// Mitsubishi GX Works2 project: AVRInfacomV3   PLC: FX3G

TYPE CutCard : STRUCT
  Lenth : DINT;
  Qnt : DINT;
END_STRUCT END_TYPE

// global labels: _io
VAR_GLOBAL
  DI_Avar1 AT X000 : BOOL;
  DI_Line1IsOff AT X001 : BOOL;
  DI_Avar2 AT X002 : BOOL;
  DI_Line2IsOff AT X003 : BOOL;
  DI_AvarGenerator AT X004 : BOOL;
  DI_GeneratorIsOff AT X005 : BOOL;
  DI_AvarSection AT X006 : BOOL;
  DI_SectionIsOff AT X007 : BOOL;
  DI_RKF1 AT X010 : BOOL;
  DI_RKF2 AT X011 : BOOL;
  DI_RKF3 AT X012 : BOOL;
  DI_Avarkontrol AT X013 : BOOL;
  DO_On1 AT Y000 : BOOL;
  DO_Off1 AT Y001 : BOOL;
  DO_On2 AT Y002 : BOOL;
  DO_Off2 AT Y003 : BOOL;
  DO_OnGenerator AT Y004 : BOOL;
  DO_OffGenerator AT Y005 : BOOL;
  DO_OnSection AT Y006 : BOOL;
  DO_OffSection AT Y007 : BOOL;
  DO_StartGenerator AT Y010 : BOOL;
END_VAR

// global labels: _gvl
VAR_GLOBAL
  gxAvto AT M400 : BOOL;
  gxOn1 AT M100 : BOOL;
  gxOff1 AT M101 : BOOL;
  gxOn2 AT M102 : BOOL;
  clTimeGenerator AT D1000 : INT;
  clTimeRKF1 AT D1001 : INT;
  clTimeRKF2 AT D1002 : INT;
  clTimeRKF3 AT D1003 : INT;
  gxOff2 AT M103 : BOOL;
  gxOnGenerator AT M104 : BOOL;
  gxOffGenerator AT M105 : BOOL;
  gxOnSection AT M106 : BOOL;
  gxOffSection AT M107 : BOOL;
  gxStartGenerator AT M108 : BOOL;
  clStartgenerator AT D1004 : INT;
  gxIsAlarm AT M150 : BOOL;
  VVALine1 : VVA;
  VVALine2 : VVA;
  VVAGen : VVA;
  VVASec : VVA;
  clTimeBackAuto AT D1005 : INT;
  gxVVAOff AT M401 : BOOL;
  gxProblemVVA1 AT M110 : BOOL;
  gxProblemVVA2 AT M111 : BOOL;
  gxProblemVVAgen AT M112 : BOOL;
END_VAR

// task Task_init (event M8002, interval 0, priority 1): PRG_INIT
// task Task_Main (event TRUE, interval 0, priority 31): POU_01
// task Task_Process (event TRUE, interval 0, priority 31): PRG_PROCESS
// user libraries (not included): AlarmManger128, Modbusv16, TimeControl, Utils

PROGRAM POU_01
VAR
  fbAmBlock : AM_IS_BLOCK;
  iStep : INT;
  wTimeRKFs : INT;
  xGenerator : BOOL;
  TPStartGen : TP;
  fbAmalarm : AM_HAS_ALARMS;
  xAllGood : BOOL;
END_VAR
(* fbAmBlock(iProcessNum := 1, iSeverity := AM_ERROR, Q := gxIsAlarm); *)
fbAmalarm(iProcessNum := 0, iSeverity := 0, Q := gxIsAlarm);
wTimeRKFs := SEL(clTimeRKF1 > clTimeRKF2, clTimeRKF2, clTimeRKF1);

IF MEF(gxAvto) THEN
    iStep := 10;
END_IF;

IF MEP(gxAvto) THEN
    iStep := 0;
END_IF;

M1 := DI_RKF1 AND NOT VVALine1.xError;
M2 := DI_RKF2 AND NOT VVALine2.xError;
M3 := DI_RKF3 AND NOT VVAGen.xError;

OUT_T(M1, TC1, SEC_TO_TIMER100(clTimeRKF1));
OUT_T(M2, TC2, SEC_TO_TIMER100(clTimeRKF2));
OUT_T(M3, TC3, SEC_TO_TIMER100(clTimeRKF3)); 

OUT_T(TRUE, TC30, 100);
OUT_T(iStep = 30 AND DI_Line1IsOff, TC4, 100);
OUT_T(iStep = 40 AND DI_Line2IsOff, TC5, 100);
OUT_T(iStep = 50 AND DI_GeneratorIsOff, TC6, 100);

(*BackAuto
OUT_T(gxVVAOff, TC31, SEC_TO_TIMER100(clTimeBackAuto));
IF TS31 THEN
	gxVVAOff := FALSE;
END_IF;
*)

CASE iStep OF
    0: (* Reset timers *)
        xGenerator := FALSE;
        gxStartGenerator := FALSE;
        MOV(TS30, 1, iStep);

    1: (* Test everything *)
    	xAllGood := TRUE;
    	
    
        MOV(xAllGood, 10, iStep);

    10: (* Idle *)

        MOV(gxAvto, 20, iStep);
        RST(gxAvto, gxStartGenerator);

		SET(
			MEP(gxOn1) 
			AND DI_Line2IsOff 
			AND DI_Line1IsOff 
			AND DI_GeneratorIsOff 
			AND DI_RKF1, 
			VVALine1.SetOn
		);
		RST( 
			MEP(gxOff1) 
			OR NOT DI_Line2IsOff 
			OR NOT DI_GeneratorIsOff 
			OR NOT DI_RKF1, 
			VVALine1.SetOn
		);

		SET(
			MEP(gxOn2) 
			AND DI_Line2IsOff 
			AND DI_Line1IsOff 
			AND DI_GeneratorIsOff 
			AND DI_RKF2, 
			VVALine2.SetOn
		);
		RST( 
			MEP(gxOff2) 
			OR NOT DI_Line1IsOff 
			OR NOT DI_GeneratorIsOff 
			OR NOT DI_RKF2, 
			VVALine2.SetOn
		);
		
		SET(
			MEP(gxOnGenerator) 
			AND DI_Line2IsOff 
			AND DI_Line1IsOff 
			AND DI_GeneratorIsOff 
			AND DI_RKF3, 
			VVAGen.SetOn
		);
		RST( 
			MEP(gxOffGenerator) 
			OR NOT DI_Line1IsOff 
			OR NOT DI_Line2IsOff 
			OR NOT DI_RKF3, 
			VVAGen.SetOn
		);
      
        xGenerator := gxStartGenerator;

    20: (* Selector *)
        MOV(TS1, 30, iStep);
        MOV(TS2 AND NOT TS1, 40, iStep);
        MOV(NOT TS1 AND NOT TS2 AND TS3, 50, iStep);
		xGenerator := NOT TS1 AND NOT TS2;

    30: (* Line 1 *)
	    VVALine2.SetOn := FALSE;
	    VVAGen.SetOn := FALSE;
        SET(TS4, gxProblemVVA1);
        SET(TS4, gxVVAOff);
        
        MOV(
        	NOT TS1 (* Контроль фаз *)
        	OR TS4 (* выключение в ручну *)
        	OR VVALine1.xError, (* автомат в ошибке *)
        	10,
        	iStep
        );

        VVALine1.SetOn := DI_GeneratorIsOff 
        	AND DI_Line2IsOff AND iStep = 30;
    
    40: (* Line 2 *)
	    VVALine1.SetOn := FALSE;
	    VVAGen.SetOn := FALSE;
        SET(TS5, gxProblemVVA2);
        SET(TS5, gxVVAOff);
         
        MOV(
        	NOT TS2 (* Контроль фаз *)
        	OR TS5 (* выключение в ручну *)
        	OR VVALine2.xError, (* автомат в ошибке *)
        	10,
        	iStep
        );

        VVALine2.SetOn := DI_GeneratorIsOff 
        	AND DI_Line1IsOff AND iStep = 40;
    
    50: (* Generator *)
	    VVALine2.SetOn := FALSE;
	    VVALine1.SetOn := FALSE;
        SET(TS6, gxProblemVVAgen);
        SET(TS6, gxVVAOff);
        
        MOV(
        	NOT TS3 (* Контроль фаз *)
        	OR TS1 OR TS2 (* появилась сеть *)
        	OR TS6 (* выключение в ручну *)
        	OR VVAGen.xError, (* автомат в ошибке *)
        	10,
        	iStep
        );
		
		xGenerator := TRUE;
        VVAGen.SetOn := DI_Line1IsOff 
        	AND DI_Line2IsOff AND iStep = 50;
END_CASE;

TPStartGen(IN := xGenerator, PT := SEC_TO_TIME(clTimeGenerator));
DO_StartGenerator := NOT (xGenerator OR TPStartGen.Q);

IF iStep > 0 THEN
	VVALine1(
		IsOn := NOT DI_Line1IsOff, 
		ResetAlarm := M2002, 
		Vkl := DO_On1, 
		Otkl := DO_Off1
	);
	VVALine2(
		IsOn := NOT DI_Line2IsOff, 
		ResetAlarm := M2002, 
		Vkl := DO_On2, 
		Otkl := DO_Off2
	);
	VVAGen(
		IsOn := NOT DI_GeneratorIsOff, 
		ResetAlarm := M2002, 
		Vkl := DO_OnGenerator, 
		Otkl := DO_OffGenerator
	);
END_IF;
END_PROGRAM

PROGRAM PRG_INIT
VAR
  fbAmInit : AM_INIT;
END_VAR
AM_D_START := 3000;

VVALine1.AlarmNum := 1;
VVALine2.AlarmNum := 2;
VVAGen.AlarmNum := 3;
VVASec.AlarmNum := 4;

(* Ошибка UPS *)
fbAmInit(iNum := 0, iSeverity := 3, iProcess := 1, xLatch := 0, xBuzzer := 0, xLock := 0);
(* Ошибка ВА Сеть 1 *)
fbAmInit(iNum := 1 , xLatch := 1, xLock := 0 );
(* Ошибка ВА Сеть 2 *)
fbAmInit(iNum := 2 , xLatch := 1, xLock := 0 );
(* Ошибка ВА Генератор *)
fbAmInit(iNum := 3 , xLatch := 1, xLock := 0 );
(* Ошибка ВА Секционный *)
fbAmInit(iNum := 4 , xLatch := 1, xLock := 0);
(* Отказ вкл ВА Сеть 1 *)
fbAmInit(iNum := 5, xLatch := 0, xLock := 0);
(* Отказ выкл ВА Сеть 1 *)
fbAmInit(iNum := 6 , xLatch := 0, xLock := 0 );
(* Отказ вкл ВА Сеть 2 *)
fbAmInit(iNum := 7 , xLatch := 0, xLock := 0 );
(* Отказ выкл ВА Сеть 2 *)
fbAmInit(iNum := 8 , xLatch := 0, xLock := 0 );
(* Отказ вкл ВА Генератор *)
fbAmInit(iNum := 9 , xLatch := 0, xLock := 0);
(* Отказ выкл ВА Генератор *)
fbAmInit(iNum := 10, xLatch := 0, xLock := 0);
(* Отказ вкл ВА Секционный *)
fbAmInit(iNum := 11 , xLatch := 0, xLock := 0 );
(* Отказ выкл ВА Секционный *)
fbAmInit(iNum := 12 , xLatch := 0, xLock := 0 );
(* Отказ запуска генератора *)
fbAmInit(iNum := 13 , xLatch := 1, xLock := 0 );
(* Данные не заполнены *)
fbAmInit(iNum := 14 , xLatch := 0, xLock := 1);
END_PROGRAM

PROGRAM PRG_PROCESS
VAR
  fbAmSet : AM_SET;
  fbAmReset : AM_RST;
  xNodata : BOOL;
  fbAMEvents : AM_EVENT;
  fbTOFResetProblems : TOF;
  PortSettings : DWORD;
  xMBInit : BOOL;
END_VAR
fbAmReset(IN := M2002);

IF  M2002 THEN
	gxProblemVVA1 := FALSE;
	gxProblemVVA2 := FALSE;
	gxProblemVVAgen := FALSE;
END_IF;

PortSettings := MB_PORT_SETTINGS(MB_PARITY_NONE, MB_STOPBIT_1, MB_BPS_38400);
xMBInit :=  MB_SLAVE_INIT_PORT2(TRUE, 20, PortSettings);

(* Тревоги *)
OUT_T(NOT DI_Avarkontrol, TC24, 10);
fbAmSet(iNum := 0, xState := TS24);
OUT_T(NOT DI_Avar1 OR gxProblemVVA1, TC21, 5);
fbAmSet(iNum := 1, xState := TS21);
OUT_T(NOT DI_Avar2 OR gxProblemVVA2, TC22, 5);
fbAmSet(iNum := 2, xState := TS22);
OUT_T(NOT DI_AvarGenerator OR gxProblemVVAgen, TC23, 5);
fbAmSet(iNum := 3, xState := TS23);
fbAmSet(iNum := 4, xState := FALSE);
OUT_T(DO_On1 AND DI_Line1IsOff, TC11, 10);
fbAmSet(iNum := 5, xState := TS11);
OUT_T(DO_Off1 AND NOT DI_Line1IsOff, TC12, 10);
fbAmSet(iNum := 6, xState := TS12);
OUT_T(DO_On2 AND DI_Line2IsOff, TC13, 10);
fbAmSet(iNum := 7, xState := TS13);
OUT_T(DO_Off2 AND NOT DI_Line2IsOff, TC14, 10);
fbAmSet(iNum := 8, xState := TS14);
OUT_T(DO_Ongenerator AND DI_GeneratorIsOff, TC15, 10);
fbAmSet(iNum := 9, xState := TS15);
OUT_T(DO_OffGenerator AND NOT DI_GeneratorIsOff, TC16, 10);
fbAmSet(iNum := 10, xState := TS16);
OUT_T(DO_OnSection AND DI_SectionIsOff , TC17, 10);
fbAmSet(iNum := 1, xState := TS17);
OUT_T(DO_OffSection AND NOT DI_SectionIsOff, TC18, 10);
fbAmSet(iNum := 12, xState := TS18);
OUT_T(NOT DO_StartGenerator AND NOT DI_RKF3, TC19, SEC_TO_TIMER100(clStartgenerator));
fbAmSet(iNum := 13, xState := TS19);

xNodata := (
	clStartgenerator = 0 
	OR clTimeGenerator = 0 
	OR clTimeRKF1 = 0 
	OR clTimeRKF2 = 0 
	OR clTimeRKF3 = 0
);
fbAmSet(iNum := 14, xState := xNodata);

fbAMEvents(EventNum := 0, EventState := DI_RKF1);
fbAMEvents(EventNum := 1, EventState := NOT DI_RKF1);
fbAMEvents(EventNum := 2, EventState := DI_RKF2);
fbAMEvents(EventNum := 3, EventState := NOT DI_RKF2);
fbAMEvents(EventNum := 4, EventState := DI_RKF3);
fbAMEvents(EventNum := 5, EventState := NOT DI_RKF3);
fbAMEvents(EventNum := 6, EventState := DO_On1);
fbAMEvents(EventNum := 7, EventState := DO_Off1);
fbAMEvents(EventNum := 8, EventState := DO_On2);
fbAMEvents(EventNum := 9, EventState := DO_Off2);
fbAMEvents(EventNum := 10, EventState := DO_Ongenerator);
fbAMEvents(EventNum := 11, EventState := DO_Offgenerator);
fbAMEvents(EventNum := 12, EventState := DO_OnSection);
fbAMEvents(EventNum := 13, EventState := DO_OffSection);
fbAMEvents(EventNum := 14, EventState := NOT DO_StartGenerator);
fbAMEvents(EventNum := 15, EventState := DO_StartGenerator);
fbAMEvents(EventNum := 16, EventState := gxAvto);
fbAMEvents(EventNum := 17, EventState := NOT gxAvto);
fbAMEvents(EventNum := 18, EventState := TS1);
fbAMEvents(EventNum := 19, EventState := TS2);
fbAMEvents(EventNum := 20, EventState := TS3);

(*
fbTOFResetProblems(IN:= MEP(gxProblemVVA1) OR MEP(gxProblemVVA2) OR MEP(gxProblemVVAgen), PT:= SEC_TO_TIME(1800));
IF  M2002 OR fbTOFResetProblems.Q THEN
	gxProblemVVA1 := FALSE;
	gxProblemVVA2 := FALSE;
	gxProblemVVAgen := FALSE;
END_IF;
*)
END_PROGRAM

FUNCTION_BLOCK VVA
VAR_IN_OUT
  SetOn : BOOL;
END_VAR
VAR_INPUT
  ResetAlarm : BOOL;
  AlarmNum : INT;
  IsOn : BOOL;
END_VAR
VAR_OUTPUT
  Vkl : BOOL;
  Otkl : BOOL;
END_VAR
VAR
  fbAmIsOn : AM_ORISON;
END_VAR
VAR_OUTPUT
  xError : BOOL;
END_VAR
VAR
  fbTPLoadBlock : TP;
  xOn : BOOL;
  xOff : BOOL;
  fbBlinkOn : BLINK;
  fbBlinkOff : BLINK;
  fbTONOn : TON;
  fbTONOff : TON;
  xTempError : BOOL;
  fbTPTON : TON;
END_VAR
RST(xError AND ResetAlarm, xError);

(* Самостоятельно октлючился в авто режиме
или сработало аварийное отключение *)
xTempError := FALSE;
fbAmIsOn(iNum := AlarmNum, Q := xTempError);

SET(fbAmIsOn.Q, xError);
SET(xError AND ResetAlarm, xOff);

fbTONOn(IN:=isOn, PT:=T#100ms);
fbTONOff(IN:=NOT isOn, PT:=T#100ms);

IF NOT xError THEN
	(* Задача включить автомат *)
	SET(MEP(SetOn) AND NOT IsOn, xOn);
	
	(* Задача отключить автомат *)
    SET(MEF(SetOn) AND IsOn, xOff);

	(* Автомат сам отключился *)
	RST(SetOn AND MEP(fbTONOff.Q), SetOn);
    
	(* Автомат сам включился *)
	RST(NOT SetOn AND MEP(fbTONOn.Q), gxAvto);
	SET(NOT SetOn AND MEP(fbTONOn.Q), SetOn);
END_IF;

(* ??? Check when spring loading *)
fbTPTON(IN:= Vkl ,PT:= T#900ms);
fbTPLoadBlock(IN := fbTPTON.Q, PT:= T#5s);

RST(MEP(xOn) OR xError, xOff);
RST(MEP(xOff) OR xError, xOn);
RST(xOn AND IsOn, xOn);
RST(xOff AND NOT IsOn, xOff);

fbBlinkOn(IN := xOn AND NOT fbTPLoadBlock.Q, 
TIMELOW:=T#1000ms, TIMEHIGH:=T#1000ms, Q := Vkl);
fbBlinkOff(IN := xOff AND NOT fbTPLoadBlock.Q, 
TIMELOW:=T#1000ms, TIMEHIGH:=T#1000ms, Q := Otkl);
END_FUNCTION_BLOCK
